(* IEC 61131-3 sources: bcs-engineering-dsl/language/test/generating/struct_test/expected, 4 files *)

(* ---- Circle.st ---- *)
TYPE Circle :
STRUCT
    radius : REAL;
END_STRUCT
END_TYPE

(* ---- Point.st ---- *)
TYPE Point :
STRUCT
    x : REAL;
    y : REAL;
END_STRUCT
END_TYPE

(* ---- Rectangle.st ---- *)
TYPE Rectangle :
STRUCT
    x : REAL;
    y : REAL;
END_STRUCT
END_TYPE

(* ---- MAIN_decl.st ---- *)
PROGRAM MAIN
VAR
    windowContact_value AT %I*: BOOL; (* Input channel from hardware *)
    TestStructs_rect: Rectangle := (x:=5, y:=10);
    TestStructs_area: REAL;
    TestStructs_perimeter: REAL;
    TestStructs_rects: ARRAY [0..1] OF Rectangle := [(x:=1, y:=2), (x:=3, y:=4)];
    TestStructs_area2: REAL := TestStructs_rects[0].x * TestStructs_rects[0].y;
END_VAR
